Staubli VAL3: safeCheck.pjx

--- safeCheck.pjx ---
Parameters version=s8.10.3Cs9_BS2093 stackSize=5000 millimeterUnit=true
Program file=computeSPoint.pgx
Program file=computeZone.pgx
Program file=iolink.pgx
Program file=loadSAFE.pgx
Program file=main.pgx
Program file=safePointCheck.pgx
Program file=safeZoneCheck.pgx
Program file=setZoneFrame.pgx
Program file=start.pgx
Program file=stop.pgx
Data file=safeCheck.dtx
Library alias=safeTemp path=Disk://source/template/safeTemp/safeTemp.pjx
Library alias=savedata path=Disk://source/saveData/saveData.pjx
Library alias=io path=Disk://source/projectSource/io/io.pjx

--- safeCheck.dtx ---
mdesc mNomSpeed
num nToolIndex
public num nIO_Zoneindex[16]
public num nIO_spindex[16]
public dio O_safePoint[16]
public dio O_safeZone

--- main.pgx ---
public program main()
begin
  //start
  call iolink()

  //main loop
  do
    call safePointCheck()


    call safeZoneCheck()


    delay(0)
  until false
end

--- start.pgx ---
program start()
begin
end

--- computeSPoint.pgx ---
public program computeSPoint(num x_nIndex, bool& x_bResult)
  local tool l_tTool
  local pointRx l_pHere
  local trsf l_trsf
  local num l_nDistance
begin
  //link(l_tTool,flange)
  //call savedata:getTool(nToolIndex,l_tTool)
  l_pHere=here(flange,world)
  l_trsf=safeTemp:sSPoint[x_nIndex].pPointRx.trsf
  l_nDistance=distance(l_pHere.trsf,l_trsf)
  if abs(l_nDistance)<5
    x_bResult=true
  else
    x_bResult=false
  endIf
end

--- computeZone.pgx ---
public program computeZone(num x_nIndex, bool& x_bResult)
  local tool l_tTool
  local frame l_fFrame
  local trsf l_trFirst
  local trsf l_trSecond
  local num l_nMax_x
  local num l_nMax_y
  local num l_nMax_z
  local num l_nMin_x
  local num l_nMin_y
  local num l_nMin_z
  local pointRx l_pPoint
  local bool l_bReuslt1
  local bool l_bReuslt2
  local bool l_bReuslt3
begin
  link(l_tTool,flange)
  link(l_fFrame,world)
  l_fFrame.trsf=safeTemp:zZoneItem[x_nIndex].fBase.trsf
  call savedata:getTool(nToolIndex,l_tTool)
  l_pPoint=here(l_tTool,l_fFrame)
  l_trFirst=safeTemp:zZoneItem[x_nIndex].pFirst.trsf
  l_trSecond=safeTemp:zZoneItem[x_nIndex].pSecond.trsf

  l_nMax_x=max(l_trFirst.x,l_trSecond.x)
  l_nMax_y=max(l_trFirst.y,l_trSecond.y)
  l_nMax_z=max(l_trFirst.z,l_trSecond.z)
  l_nMin_x=min(l_trFirst.x,l_trSecond.x)
  l_nMin_y=min(l_trFirst.y,l_trSecond.y)
  l_nMin_z=min(l_trFirst.z,l_trSecond.z)

  if l_nMin_x<l_pPoint.trsf.x and l_pPoint.trsf.x<l_nMax_x
    l_bReuslt1=true
  else
    l_bReuslt1=false
  endIf

  if l_nMin_y<l_pPoint.trsf.y and l_pPoint.trsf.y<l_nMax_y
    l_bReuslt2=true
  else
    l_bReuslt2=false
  endIf

  if l_nMin_z<l_pPoint.trsf.z and l_pPoint.trsf.z<l_nMax_z
    l_bReuslt3=true
  else
    l_bReuslt3=false
  endIf

  if l_bReuslt1 and l_bReuslt2 and l_bReuslt3
    x_bResult=true
  else
    x_bResult=false
  endIf
end

--- iolink.pgx ---
public program iolink()
  local num l_i
begin
  for l_i = 0 to size(O_safePoint)-1
    dioLink(O_safePoint[l_i],io:dOutput[nIO_spindex[l_i]])
  endFor

  for l_i =0 to size(O_safeZone)-1
    dioLink(O_safeZone[l_i],io:dOutput[nIO_Zoneindex[l_i]])
  endFor
end

--- loadSAFE.pgx ---
public program loadSAFE(num x_nLib, num& x_nResult)
  local string l_sPath
begin
  l_sPath="Disk://data/CustomerLib/lib"+toString("",x_nLib)+"/safeData/safeData.pjx"
  x_nResult=safeTemp:libLoad(l_sPath)
  delay(0)
  logMsg(toString("",x_nResult))
end

--- safePointCheck.pgx ---
public program safePointCheck()
  local bool l_bResult
  local bool l_bErr
  local num l_i
begin
  for l_i = 0 to size(safeTemp:sSPoint)-1
    call computeSPoint(l_i,l_bResult)
    //O_safePoint[l_i]=(l_bResult==true)
    call io:setDigOutput(O_safePoint[l_i],l_bResult,l_bErr)
  endFor
end

--- safeZoneCheck.pgx ---
public program safeZoneCheck()
  local bool l_bResult
  local bool l_bErr
  local num l_i
begin
  for l_i = 0 to size(safeTemp:zZoneItem)-1
    if safeTemp:zZoneItem[l_i].bActive
      call computeZone(l_i,l_bResult)
      call io:setDigOutput(O_safeZone[l_i],l_bResult,l_bErr)
    endIf
  endFor
end

--- setZoneFrame.pgx ---
public program setZoneFrame()
  local num x_nIndex
  local pointRx l_pPoint1
  local pointRx l_pPoint2
  local pointRx l_pPoint3
  local num l_nResult
begin
  link(l_pPoint1,world)
  link(l_pPoint2,world)
  link(l_pPoint3,world)
  l_pPoint1=safeTemp:zZoneItem[x_nIndex].pO
  l_pPoint2=safeTemp:zZoneItem[x_nIndex].pX
  l_pPoint3=safeTemp:zZoneItem[x_nIndex].pY
  l_nResult=setFrame(l_pPoint1,l_pPoint2,l_pPoint3,safeTemp:zZoneItem[x_nIndex].fBase)
  if l_nResult<0
    userPageAlert("坐标系生成失败："+toString("",x_nIndex))
    logMsg("坐标系生成失败："+toString("",x_nIndex))
  endIf
end

--- stop.pgx ---
program stop()
begin
end
